Universal Robots PolyScope program: TgtProg.urp

Program TgtProg (createdIn=3.0.0 lastSavedIn=3.0.0 directory=/programs installation=default)
Robot Program (runOnlyOnce=true motionType=MoveJ speed=1.047198 acceleration=1.396263 useActiveTCP=false)
  'Program generated by RoboDK v6.0.7 for UR10 on XX/XX/XXXX 18:00:00'
  'Using nominal kinematics.'
  Set DigitalOutput pin=digital_out[12]; digitalValue=1
  Set DigitalOutput pin=digital_out[25]; digitalValue=true
  Set DigitalOutput pin=digital_out[3]; digitalValue=False
  Set DigitalOutput pin=digital_out[4]; digitalValue=0
  Wait DigitalInput pin=digital_in[get_standard_digital_in(15)]; digitalValue=1
  Wait DigitalInput pin=digital_in[get_standard_digital_in(22)]; digitalValue=off
  Set DigitalOutput pin=digital_out[2]; digitalValue=1
  Set DigitalOutput pin=digital_out[5]; digitalValue=0
  Call Call_A
  Call Call_B
  Call Call_A
SubProgram  [hidden by the author, left out]
SubProgram  [hidden by the author, left out]
SubProgram Call_A [hidden by the author, left out]
SubProgram Call_B [hidden by the author, left out]
